(* IEC 61131-3 sources: daoli-st-library/DL_Device (part 39) *)

(* ---- FB_DL_HeatCoolZone.st ---- *)
(*==============================================================================
 * 组件名称 (Component)  : FB_DL_HeatCoolZone
 * 所属子库 (Sublibrary) : DL_Device
 * 当前版本 (Version)    : 1.0.0
 * 兼容性   (Platform)   : CODESYS 3.5 / TwinCAT 3 / 汇川 InoProShop / Machine Expert
 *                         仅依赖 Standard.library 语义与 DL_Algo 既有算法组件，
 *                         零厂商方言，零物理地址直写
 * 分类     (Category)   : 功能块（FUNCTION_BLOCK）· 加热/冷却温控区 · Level 1 DL_Device 开库件
 * 功能描述 (Function)   : 双通道（加热/冷却）温控区控制器，R4 算法族首个上层消费者。
 *                         控制链：FB_DL_PidController（含抗饱和，实例经引脚注入，
 *                         参数外置组态）→ 分程分配（Split-range，fSplitLow/High
 *                         可组态，非魔法数）→ FB_DL_PwmDutyController × 2（加热/
 *                         冷却 SSR 驱动）。断偶保护：传感器接口信号质量进入断线/
 *                         开路域时按 eBreakAction 切断对应通道并锁存 eSensorBreak
 *                         态（0003_0211），退出需 CmdReset 且质量恢复 eGood；
 *                         锁存期间双通道全断为最终安全态。设定值经 fTempMin/Max
 *                         钳位（信息级 0003_0101，不置故障）。本块零内嵌组态、
 *                         零魔法数，PID/PWM 全部实例经 IN_OUT 引脚注入。
 * 开源溯源 (Origin)     : 原创实现。分程控制与断偶安全方向为行业公知语义
 *                         （来源标签 lbp-device；断偶方向参考 NAMUR NE43 公开
 *                         标准），未复制任何厂商源码。PID/PWM 语义消费本库
 *                         DL_Algo 既有组件 FB_DL_PidController / FB_DL_PwmDutyController。
 * 本文件内含       : TYPE      E_DL_BreakAction（断偶动作方向枚举，归属 DL_Device）
 *                    FUNCTION_BLOCK FB_DL_HeatCoolZone IMPLEMENTS I_DL_TemperatureZone
 *                    （随附 METHOD ×3 与 PROPERTY GET ×5 实现体）
 * 依赖     (Depends)    : I_DL_TemperatureZone / E_DL_TempZoneState（同轮泳道交付
 *                          的 I_DL_TemperatureZone.st）；FB_DL_PidController、
 *                          FB_DL_PwmDutyController（DL_Algo v1.0.1+，实例注入）；
 *                          Standard.library：LIMIT / MIN / ABS。不引用库内任何
 *                          其他实现文件的具体逻辑。
 * 【规格偏离留档 / R11 Deviation register】
 *   D1 规格 §1.8 引脚表要求 fTempActual/fPowerOut/eState/bFault/uErrorId 五个
 *      「接口属性映射」成员同时作为 OUT 引脚暴露；IEC 61131-3 同一 POU 的变量
 *      与属性共享命名空间，同名变量与同名属性并存无法通过编译。按 R11 留档：
 *      该五成员以只读 PROPERTY 形式对外暴露（属性即输出引脚语义，接口成员逐一
 *      兑现），bHeaterOut/bCoolerOut 两个非接口成员保留 VAR_OUTPUT。
 *   D2（已闭环 / Closed）规格 §1.5 的 E_DL_SignalQuality / I_DL_AnalogSensor 为
 *      本块温度信号源契约。编码阶段宿主文件未入库，本文件曾就地声明副本；
 *      R5 注册收口阶段 I_DL_AnalogSensor.st（正式承载 E_DL_SignalQuality 枚举
 *      与 I_DL_AnalogSensor 接口）已随 DL_Device 开库交付，本文件重复副本已
 *      删除，改为引用该正式定义（IEC 同工程内 INTERFACE/ENUM 全局可见，与原
 *      D2 预设处置一致）。契约语义以 I_DL_AnalogSensor.st 为准（本块仅消费
 *      fValue 与 eQuality 两个成员）。
 *   D3 规格 §1.8「按 eBreakAction 切断对应通道并锁存」细化：eBreakAction 决定
 *      断偶瞬间立即切断的危险通道方向；锁存 eSensorBreak 期间双通道全断为最终
 *      安全态（锁存态不维持任何输出，安全侧选择）。
 *   D4 公约 0.6 示例码 16#0001_0001 属 DL_Base 段；按公约 0.7 段位分配（DL_Device
 *      族 16#0003_xxxx），本块参数钳位/对调修复统一置信息级 16#0003_0101。
 *   D5 新增故障/信息码顺延登记（无冲突）：16#0003_0212 非法状态兜底（故障级）、
 *      16#0003_0213 传感器接口引用未注入/无效（故障级）。
 * 故障码表（本块全部登记，0=无故障）：
 *   16#0003_0101【信息级】参数钳位/对调修复/设定值钳位提示，不置故障
 *   16#0003_0211【故障级】传感器断线/开路锁存，CmdReset + 质量恢复 eGood 方可清
 *   16#0003_0212【故障级】非法状态兜底（CASE ELSE 落点），CmdReset 可清
 *   16#0003_0213【故障级】温度传感器接口引用未注入/无效，CmdReset + 引脚有效方可清
 * 红线自检 (Redline)    : R1 ✓ 零全局变量表与外部变量引用 ｜ R2 ✓ 零物理 IO 地址直写
 *                         R3 ✓ 纯 IEC 61131-3 ｜ R4 ✓ 防除零+钳位+非有限值防御+浮点容差
 *                         R5 ✓ 全变量中英双语同行注释 ｜ R6 ✓ 六态 ENUM+CASE+ELSE 兜底
 *                         R7 ✓ 无直接定时器实例（PID/PWM 实例每拍无条件调用）
 * 修订历史 (Revision)   :
 *   2026-11-15  v1.0.0  首版入库 · Round 05 · 泳道 B · 契约出处 ROUND_PLAN_R5 §1.8
 *   2026-11-15  v1.0.0  R5 收口：删除就地重复的 E_DL_SignalQuality /
 *                       I_DL_AnalogSensor 声明，改引用 I_DL_AnalogSensor.st
 *                       正式定义（D2 闭环），功能与引脚零变更
 * 验收向量 (Acceptance) :
 *   V1 正常跃迁链：bEnable=TRUE → eHolding；fTempActual 低于设定 → eHeating；
 *      回到中性带 → eHolding；高于设定 → eCooling（fPowerOut 正负号随之翻转）
 *   V2 非法态兜底：强写内部状态为越界值 → CASE ELSE 落入 eFault（0003_0212）
 *   V3 中途跟踪脉冲（公约 0.1 必含）：闭环运行中 bTrack 单拍脉冲 + fTrackValue
 *      =30.0 → 本拍 PID 输出跟随 30.0，双通道占空比无扰重分配，无输出踢腿
 *   V4 断偶：eQuality=eWireBreakHigh → 按 eBreakAction 切断并锁存 eSensorBreak
 *      （0003_0211）；质量恢复 eGood + CmdReset → 回 eHolding（带无扰同步）
 *   V5 设定值钳位：fTempSetpoint=500 且 fTempMax=300 → 生效 300，0003_0101，
 *      故障位保持 FALSE（R21 信息级不置故障）
 *   V6 参数对调：fTempMin=300 > fTempMax=0 → 对调后继续计算，0003_0101
 *   V7 引脚无效：iTempSensor 未注入 → eFault（0003_0213），双通道切断
 *============================================================================*)

(*-----------------------------------------------------------------------------
 * 契约引用说明（R5 收口）: 本块温度信号源契约 E_DL_SignalQuality 与
 * I_DL_AnalogSensor 不在本文件就地声明，统一引用 DL_Device 正式定义文件
 * I_DL_AnalogSensor.st（枚举随宿主接口文件同文件发布，IEC 同工程内全局可见，
 * 留档见头注释 D2）。本块仅消费 fValue 与 eQuality 两个成员。
 *----------------------------------------------------------------------------*)

(*-----------------------------------------------------------------------------
 * 枚举: E_DL_BreakAction（归属 DL_Device，随 FB_DL_HeatCoolZone 同文件）
 * 含义: 断偶动作方向，按被控对象安全策略配置。
 *----------------------------------------------------------------------------*)
{attribute 'qualified_only'}
{attribute 'strict'}
TYPE E_DL_BreakAction :
(
    eHeatOff := 0,   // 断偶切断加热（Cut heating on break）：升温对象超温风险侧
    eCoolOff := 1    // 断偶切断冷却（Cut cooling on break）：骤冷风险对象（如防脆断工艺）侧
) UINT;
END_TYPE

(*==============================================================================
 * 功能块: FB_DL_HeatCoolZone IMPLEMENTS I_DL_TemperatureZone
 * 调用约定: 每个扫描周期无条件调用一次；PID/PWM 注入实例在本块主体每拍无条件
 *           调用（不在任何 IF/CASE 分支内部）；方法仅置请求标志，动作由主体执行。
 * 分程约定: PID 输出 [0..100 %]。输出低于 fSplitLow → 加热段（越低加热越强，
 *           配合 fKp 负值反作用）；高于 fSplitHigh → 冷却段（越高冷却越强）；
 *           两点之间为中性带（双通道全关，热平衡保持）。fSplitLow=0 时加热段
 *           跨度为零、加热通道自动禁用（防除零）；fSplitHigh=100 时同理禁用冷却。
 *============================================================================*)
FUNCTION_BLOCK FB_DL_HeatCoolZone IMPLEMENTS I_DL_TemperatureZone
VAR_INPUT
    fTempSetpoint   : REAL := 0.0;      // 目标温度（Setpoint）[°C]，经 fTempMin/Max 钳位后生效
    fTempMin        : REAL := 0.0;     // 设定值下边界（Setpoint lower bound）[°C]，默认 0.0
    fTempMax        : REAL := 300.0;   // 设定值上边界（Setpoint upper bound）[°C]，默认 300.0
    fSplitLow       : REAL := 50.0;    // 分程下切换点（Split-range low crossover）[%]，PID 输出低于此点进入加热段
    fSplitHigh      : REAL := 50.0;    // 分程上切换点（Split-range high crossover）[%]，PID 输出高于此点进入冷却段
    eBreakAction    : E_DL_BreakAction := E_DL_BreakAction.eHeatOff; // 断偶动作方向（Break action）：eHeatOff=切断加热 / eCoolOff=切断冷却
    bEnable         : BOOL := FALSE;   // 投运使能（Zone enable），与 CmdEnable 方法锁存值取与
    tSampleTime     : TIME := T#100MS; // 采样周期（Sample time），下传注入的 PID 与两路 PWM（公约 0.5）
    bTrack          : BOOL := FALSE;   // 跟踪使能（Track enable），TRUE 时本拍输出跟随 fTrackValue 无扰接管
    fTrackValue     : REAL := 0.0;     // 跟踪值（Track value）[-100..100 %]，与输出功率同量纲
END_VAR
VAR_IN_OUT
    iTempSensor     : I_DL_AnalogSensor;       // 温度信号源接口引用（Sensor interface reference），上层注入 FB_DL_AnalogTransmitter 实例
    fbPid           : FB_DL_PidController;     // 温度 PID 实例（Injected PID instance），增益/积分/限幅由调用方组态
    fbPwmHeat       : FB_DL_PwmDutyController; // 加热 SSR PWM 实例（Injected heat PWM），周期/最短脉冲由调用方组态
    fbPwmCool       : FB_DL_PwmDutyController; // 冷却 SSR PWM 实例（Injected cool PWM），周期/最短脉冲由调用方组态
END_VAR
VAR_OUTPUT
    bHeaterOut      : BOOL;            // 加热执行通道镜像（Heater channel mirror），等于加热 PWM 实例布尔输出
    bCoolerOut      : BOOL;            // 冷却执行通道镜像（Cooler channel mirror），等于冷却 PWM 实例布尔输出
END_VAR
VAR
    bInit           : BOOL := TRUE;    // 首扫标志（First-scan flag），首扫判据见段 1（公约 0.1 唯一合法范式）
    _eState         : E_DL_TempZoneState := E_DL_TempZoneState.eIdle; // 内部状态机步序（Internal zone state）
    _fTempActual    : REAL := 0.0;     // 实测温度快照（Actual temperature snapshot）[°C]，取自传感器接口
    _fPowerOut      : REAL := 0.0;     // 输出功率（Power output）[-100..100 %]，正=加热 / 负=冷却（R20 量纲与赋值式一致）
    _bFault         : BOOL := FALSE;   // 故障锁存标志（Fault latched），派生式：仅故障级状态置位，信息级不置位（R21）
    _uErrorId       : UDINT := 0;      // 故障/信息码（Error/info code），0=无；故障级进态写入、锁存保持
    _bCmdEnabled    : BOOL := TRUE;    // CmdEnable 方法锁存值（Method enable latch），默认投运（方法为可选入口）
    _fSetpointMethod: REAL := 0.0;     // SetSetpoint 方法锁存设定值（Method setpoint latch）[°C]，已按边界钳位
    _bUseMethodSp   : BOOL := FALSE;   // TRUE=方法设定值覆盖引脚设定值（Method setpoint override）
    _bSyncReq       : BOOL := FALSE;   // 跃迁无扰同步请求（Bumpless sync request），置位后下一拍 PID 跟踪当前功率
    _bTrackActive   : BOOL := FALSE;   // 本拍处于外部跟踪（External track active this scan），由段 1 判据得出
    _fPowerOutLast  : REAL := 0.0;     // 上一拍输出功率（Last power output）[-100..100 %]，跃迁同步的跟踪源
    _fTempMinEff    : REAL := 0.0;     // 修复后设定值下边界（Repaired lower bound）[°C]
    _fTempMaxEff    : REAL := 300.0;   // 修复后设定值上边界（Repaired upper bound）[°C]
    _fSplitLowEff   : REAL := 50.0;    // 修复后分程下切换点（Repaired low crossover）[%]
    _fSplitHighEff  : REAL := 50.0;    // 修复后分程上切换点（Repaired high crossover）[%]
    _fSpEff         : REAL := 0.0;     // 有效设定值（Effective setpoint）[°C]，来源仲裁 + 钳位后
    _fTrackSrc      : REAL := 0.0;     // 本拍跟踪源（Track source this scan）[-100..100 %]
    _fPidOut        : REAL := 0.0;     // PID 输出快照（PID output snapshot）[0..100 %]
    _fHeatDuty      : REAL := 0.0;     // 加热通道占空比（Heater duty）[0..100 %]
    _fCoolDuty      : REAL := 0.0;     // 冷却通道占空比（Cooler duty）[0..100 %]
    _fSpTmp         : REAL := 0.0;     // 参数对调临时变量（Swap temporary）[°C 或 %]
    _bRefOk         : BOOL := FALSE;   // 传感器接口引用有效标志（Sensor reference valid）
    _bSensorBad     : BOOL := FALSE;   // 传感器断线/开路标志（Sensor break flag），含非有限值防御归入
    _bInfoClamp     : BOOL := FALSE;   // 本拍发生钳位/对调修复（Info-level clamp occurred）
    _bRunPre        : BOOL := FALSE;   // CASE 前运行态判定（Pre-CASE running flag），PID 使能源
    _bZoneRun       : BOOL := FALSE;   // CASE 后运行态判定（Post-CASE running flag），PWM 使能源
    _bReqEnable     : BOOL := FALSE;   // CmdEnable 请求挂起（Enable request pending）
    _bValEnable     : BOOL := FALSE;   // CmdEnable 请求值（Enable request value）
    _bReqReset      : BOOL := FALSE;   // CmdReset 请求挂起（Reset request pending）
    _bReqSetSp      : BOOL := FALSE;   // SetSetpoint 请求挂起（Setpoint request pending）
    _fReqSetSp      : REAL := 0.0;     // SetSetpoint 请求原始值（Raw setpoint request）[°C]
    _eQuality       : E_DL_SignalQuality := E_DL_SignalQuality.eGood; // 传感器信号质量快照（Quality snapshot）
END_VAR
VAR CONSTANT
    DL_ZONE_POWER_TOL : REAL := 0.01;   // 热平衡零功率判定容差（Power tolerance）[%]，浮点容差红线，状态判稳阈值
    DL_ZONE_SPAN_EPS  : REAL := 1.0E-6; // 分程跨度防除零判据（Span epsilon）[%]，低于此值通道禁用
END_VAR

METHOD SetSetpoint : BOOL
VAR_INPUT
    fTemp : REAL;                        // 目标温度（Target temperature）[°C]，非有限值拒绝
END_VAR
// 返回合法性：非有限值一律拒绝（公约 0.8 判式），合法值锁存待主体钳位生效
IF fTemp <> fTemp THEN
    SetSetpoint := FALSE;                // 非有限值拒绝
ELSE
    _fReqSetSp := fTemp;                 // 请求原始值 [°C]
    _bReqSetSp := TRUE;                  // 置单发标志，主体段 2/段 3 落实
    SetSetpoint := TRUE;                 // 受理成功
END_IF

    END_METHOD

METHOD CmdEnable
VAR_INPUT
    bOn : BOOL;                          // TRUE=投运（Commission on），FALSE=退出并切断双通道
END_VAR
_bReqEnable := TRUE;                     // 置请求标志
_bValEnable := bOn;                      // 请求值随行

    END_METHOD

METHOD CmdReset : BOOL
// 返回当前是否可复位：断偶锁存态要求信号质量快照已恢复 eGood（规格 §1.8 退出条件）
_bReqReset := TRUE;                      // 置请求标志，主体段 7 各态消费
IF _eState = E_DL_TempZoneState.eSensorBreak THEN
    IF _bRefOk AND (_eQuality = E_DL_SignalQuality.eGood) AND (NOT _bSensorBad) THEN
        CmdReset := TRUE;                // 质量已恢复，可复位
    ELSE
        CmdReset := FALSE;               // 仍在断线域，拒绝复位
    END_IF
ELSE
    CmdReset := TRUE;                    // 非断偶态一律受理
END_IF

// =============================================================================
// 属性实现区（PROPERTY GET ×5，接口契约逐字兑现；偏离 D1：属性即输出引脚语义）
// =============================================================================

    END_METHOD

// -----------------------------------------------------------------------------
// 段 1｜首扫与跟踪同步（公约 0.1 / R19 唯一合法范式：跟踪项在前、首扫项取反在后，
//       禁止两项顺序颠倒的反式写法；验收向量 V3 覆盖运行中途跟踪脉冲）
// -----------------------------------------------------------------------------
IF bTrack OR (NOT bInit) THEN
    _fPowerOutLast := 0.0;               // 首扫/外部跟踪：历史功率清零，杜绝接管瞬间踢腿 [±100 %]
    _bTrackActive  := TRUE;              // 本拍输出跟随外部跟踪值 fTrackValue
    bInit          := TRUE;              // 首扫完成置位
ELSE
    _bTrackActive  := FALSE;             // 正常闭环拍，跟踪源取内部历史功率
END_IF

// -----------------------------------------------------------------------------
// 段 2｜方法请求消费（方法内只置标志，动作在本周期落实——跨周期动作不驻留方法）
// -----------------------------------------------------------------------------
IF _bReqEnable THEN
    _bCmdEnabled := _bValEnable;         // 投/退锁存值更新
    _bReqEnable  := FALSE;               // 单发消费
END_IF
IF _bReqSetSp THEN
    _fSetpointMethod := _fReqSetSp;      // 方法设定值锁存 [°C]，边界钳位在段 3 统一进行
    _bUseMethodSp    := TRUE;            // 方法设定值覆盖引脚设定值
    _bReqSetSp       := FALSE;           // 单发消费
END_IF
IF NOT ( (_eState = E_DL_TempZoneState.eSensorBreak) OR (_eState = E_DL_TempZoneState.eFault) ) THEN
    _bReqReset := FALSE;                 // 非锁存态下的复位请求立即作废，防陈旧请求迟到生效
END_IF

// -----------------------------------------------------------------------------
// 段 3｜参数修复（公约 0.6 对调自修复 + 公约 0.8 非有限值防御；信息级 0003_0101
//       只进 uErrorId 不置故障，R21；偏离 D4：段位按公约 0.7 归 DL_Device 族）
// -----------------------------------------------------------------------------
_bInfoClamp := FALSE;
IF fTempMin <> fTempMin THEN             // NaN 恒不等于自身（公约 0.8 指定判式）
    _fTempMinEff := 0.0;                 // 非有限值回退默认下边界 [°C]
    _bInfoClamp  := TRUE;
ELSE
    _fTempMinEff := fTempMin;            // 直接采纳 [°C]
END_IF
IF fTempMax <> fTempMax THEN
    _fTempMaxEff := 300.0;               // 非有限值回退默认上边界 [°C]
    _bInfoClamp  := TRUE;
ELSE
    _fTempMaxEff := fTempMax;            // 直接采纳 [°C]
END_IF
IF _fTempMinEff > _fTempMaxEff THEN      // 边界对调自修复（公约 0.6）：修复后继续计算，不中断
    _fSpTmp       := _fTempMinEff;
    _fTempMinEff  := _fTempMaxEff;
    _fTempMaxEff  := _fSpTmp;
    _bInfoClamp   := TRUE;
END_IF

IF fSplitLow <> fSplitLow THEN
    _fSplitLowEff := 50.0;               // 非有限值回退对称默认 [%]
    _bInfoClamp   := TRUE;
ELSE
    _fSplitLowEff := fSplitLow;          // 直接采纳 [%]
END_IF
IF fSplitHigh <> fSplitHigh THEN
    _fSplitHighEff := 50.0;              // 非有限值回退对称默认 [%]
    _bInfoClamp    := TRUE;
ELSE
    _fSplitHighEff := fSplitHigh;        // 直接采纳 [%]
END_IF
IF _fSplitLowEff < 0.0 THEN
    _fSplitLowEff := 0.0;                // 钳到分程域下限 [%]（此时加热段跨度为零，加热禁用）
    _bInfoClamp   := TRUE;
END_IF
IF _fSplitLowEff > 100.0 THEN
    _fSplitLowEff := 100.0;              // 钳到分程域上限 [%]
    _bInfoClamp   := TRUE;
END_IF
IF _fSplitHighEff < 0.0 THEN
    _fSplitHighEff := 0.0;               // 钳到分程域下限 [%]
    _bInfoClamp    := TRUE;
END_IF
IF _fSplitHighEff > 100.0 THEN
    _fSplitHighEff := 100.0;             // 钳到分程域上限 [%]（此时冷却段跨度为零，冷却禁用）
    _bInfoClamp    := TRUE;
END_IF
IF _fSplitLowEff > _fSplitHighEff THEN   // 分程点对调自修复（公约 0.6）
    _fSpTmp        := _fSplitLowEff;
    _fSplitLowEff  := _fSplitHighEff;
    _fSplitHighEff := _fSpTmp;
    _bInfoClamp    := TRUE;
END_IF

// 设定值来源仲裁：方法锁存值优先，否则取引脚连续值
IF _bUseMethodSp THEN
    _fSpEff := _fSetpointMethod;         // 方法通道 [°C]
ELSE
    _fSpEff := fTempSetpoint;            // 引脚通道 [°C]
END_IF
IF _fSpEff <> _fSpEff THEN
    _fSpEff     := _fTempMinEff;         // 非有限设定值回退下边界（安全侧低温待机）[°C]
    _bInfoClamp := TRUE;
END_IF
IF (_fSpEff < _fTempMinEff) OR (_fSpEff > _fTempMaxEff) THEN
    _fSpEff     := LIMIT(_fTempMinEff, _fSpEff, _fTempMaxEff);  // 设定值钳位（规格 §1.8 设计点，信息级 0003_0101）
    _bInfoClamp := TRUE;
END_IF

// -----------------------------------------------------------------------------
// 段 4｜传感器采集与有效性判定（接口引用检查 + 质量域 + 非有限值防御）
// -----------------------------------------------------------------------------
_bRefOk     := FALSE;
_bSensorBad := FALSE;
_eQuality   := E_DL_SignalQuality.eGood;
IF iTempSensor <> 0 THEN                 // 接口引用有效性检查（未注入防御）
    _bRefOk     := TRUE;
    _fTempActual := iTempSensor.fValue;  // 工程量实测值 [°C]，契约保证 NaN 防御后输出
    _eQuality    := iTempSensor.eQuality;
    IF _fTempActual <> _fTempActual THEN
        _bSensorBad := TRUE;             // 非有限值防御：NaN 按断线域处理（公约 0.8 判式）
    ELSIF (_eQuality = E_DL_SignalQuality.eWireBreakLow)
       OR (_eQuality = E_DL_SignalQuality.eWireBreakHigh)
       OR (_eQuality = E_DL_SignalQuality.eOpenLoop) THEN
        _bSensorBad := TRUE;             // NE43 断线/开路域（规格 §1.8 断偶保护集合）
    END_IF
END_IF

// -----------------------------------------------------------------------------
// 段 5｜运行态预判定与注入 PID 无条件调用（R7 精神：实例调用不在 IF/CASE 分支内）
// -----------------------------------------------------------------------------
_bRunPre := (_eState = E_DL_TempZoneState.eHolding)
         OR (_eState = E_DL_TempZoneState.eHeating)
         OR (_eState = E_DL_TempZoneState.eCooling);
IF _bTrackActive THEN
    _fTrackSrc := fTrackValue;           // 外部跟踪源 [-100..100 %]
ELSE
    _fTrackSrc := _fPowerOutLast;        // 跃迁同步源 = 上一拍实际输出功率 [-100..100 %]
END_IF
fbPid(
    bEnable     := _bRunPre AND _bRefOk AND (NOT _bSensorBad),  // 断偶/无引用时冻结 PID（输出回下限）
    bManual     := FALSE,                // 温控区纯自动模式，手动路径不由本块开放
    fSetpoint   := _fSpEff,              // 有效设定值 [°C]
    fActual     := _fTempActual,         // 实测温度 [°C]
    tSampleTime := tSampleTime,          // 采样周期下传（公约 0.5）
    bTrack      := _bTrackActive OR _bSyncReq,  // 外部跟踪或跃迁无扰同步（电平，一拍）
    fTrackValue := _fTrackSrc            // 跟踪值 [-100..100 %]
);
_bSyncReq := FALSE;                      // 同步请求单发消费（段 7 跃迁时重新置位）

// -----------------------------------------------------------------------------
// 段 6｜分程分配（热平衡计算，防除零：跨度不足的通道自动禁用，R4 红线）
// -----------------------------------------------------------------------------
IF _bRunPre AND _bRefOk AND (NOT _bSensorBad) THEN
    _fPidOut := fbPid.fOut;              // PID 输出 [0..100 %]，量程由调用方组态
    IF _fPidOut < _fSplitLowEff THEN
        // 加热段：输出越低于下切换点，加热越强（配合 fKp 负值反作用惯例）
        IF _fSplitLowEff > DL_ZONE_SPAN_EPS THEN
            _fHeatDuty := LIMIT(0.0, (_fSplitLowEff - _fPidOut) / _fSplitLowEff * 100.0, 100.0); // 加热占空比 [0..100 %]
        ELSE
            _fHeatDuty := 0.0;           // 加热段跨度为零，通道禁用（防除零）
        END_IF
        _fCoolDuty := 0.0;               // 加热段冷却通道必关 [0..100 %]
    ELSIF _fPidOut > _fSplitHighEff THEN
        // 冷却段：输出越高于上切换点，冷却越强
        IF (100.0 - _fSplitHighEff) > DL_ZONE_SPAN_EPS THEN
            _fCoolDuty := LIMIT(0.0, (_fPidOut - _fSplitHighEff) / (100.0 - _fSplitHighEff) * 100.0, 100.0); // 冷却占空比 [0..100 %]
        ELSE
            _fCoolDuty := 0.0;           // 冷却段跨度为零，通道禁用（防除零）
        END_IF
        _fHeatDuty := 0.0;               // 冷却段加热通道必关 [0..100 %]
    ELSE
        _fHeatDuty := 0.0;               // 中性带：双通道全关，热平衡保持 [0..100 %]
        _fCoolDuty := 0.0;               // 中性带 [0..100 %]
    END_IF
ELSE
    _fPidOut   := 0.0;                   // 非运行拍 PID 输出按 0 [%] 处理
    _fHeatDuty := 0.0;                   // 非运行拍加热占空比清零 [0..100 %]
    _fCoolDuty := 0.0;                   // 非运行拍冷却占空比清零 [0..100 %]
END_IF
_fPowerOut := _fHeatDuty - _fCoolDuty;   // 输出功率 [-100..100 %]，正=加热/负=冷却（R20 量纲与赋值式一致）

// -----------------------------------------------------------------------------
// 段 7｜状态机（ENUM + CASE + ELSE 兜底；断偶/非法态/无引用均为锁存，R15 仅复位可清）
// -----------------------------------------------------------------------------
CASE _eState OF

    E_DL_TempZoneState.eIdle:            // 空闲：双通道切断（PWM 使能在段 8 落实）
        IF _bRefOk AND (NOT _bSensorBad) AND bEnable AND _bCmdEnabled THEN
            _bSyncReq := TRUE;           // 投运首拍无扰同步，PID 跟踪当前功率 0 [%]
            _eState   := E_DL_TempZoneState.eHolding;
        END_IF

    E_DL_TempZoneState.eHolding:         // 保温：双通道处于热平衡容差带
        IF NOT (bEnable AND _bCmdEnabled) THEN
            _eState := E_DL_TempZoneState.eIdle;
        ELSIF NOT _bRefOk THEN
            _uErrorId := 16#0003_0213;   // 接口引用未注入/无效（故障级锁存）
            _eState   := E_DL_TempZoneState.eFault;
        ELSIF _bSensorBad THEN
            _uErrorId := 16#0003_0211;   // 断偶锁存（故障级；eBreakAction 切断方向语义见偏离 D3）
            _eState   := E_DL_TempZoneState.eSensorBreak;
        ELSIF _fPowerOut > DL_ZONE_POWER_TOL THEN
            _eState := E_DL_TempZoneState.eHeating;
        ELSIF _fPowerOut < -DL_ZONE_POWER_TOL THEN
            _eState := E_DL_TempZoneState.eCooling;
        END_IF

    E_DL_TempZoneState.eHeating:         // 加热中
        IF NOT (bEnable AND _bCmdEnabled) THEN
            _eState := E_DL_TempZoneState.eIdle;
        ELSIF NOT _bRefOk THEN
            _uErrorId := 16#0003_0213;   // 接口引用未注入/无效
            _eState   := E_DL_TempZoneState.eFault;
        ELSIF _bSensorBad THEN
            _uErrorId := 16#0003_0211;   // 断偶锁存
            _eState   := E_DL_TempZoneState.eSensorBreak;
        ELSIF _fPowerOut < -DL_ZONE_POWER_TOL THEN
            _eState := E_DL_TempZoneState.eCooling;
        ELSIF ABS(_fPowerOut) <= DL_ZONE_POWER_TOL THEN
            _eState := E_DL_TempZoneState.eHolding;   // 回到热平衡带（浮点容差红线）
        END_IF

    E_DL_TempZoneState.eCooling:         // 冷却中
        IF NOT (bEnable AND _bCmdEnabled) THEN
            _eState := E_DL_TempZoneState.eIdle;
        ELSIF NOT _bRefOk THEN
            _uErrorId := 16#0003_0213;   // 接口引用未注入/无效
            _eState   := E_DL_TempZoneState.eFault;
        ELSIF _bSensorBad THEN
            _uErrorId := 16#0003_0211;   // 断偶锁存
            _eState   := E_DL_TempZoneState.eSensorBreak;
        ELSIF _fPowerOut > DL_ZONE_POWER_TOL THEN
            _eState := E_DL_TempZoneState.eHeating;
        ELSIF ABS(_fPowerOut) <= DL_ZONE_POWER_TOL THEN
            _eState := E_DL_TempZoneState.eHolding;   // 回到热平衡带
        END_IF

    E_DL_TempZoneState.eSensorBreak:     // 断偶锁存：双通道全断（安全终态，偏离 D3）
        IF _bReqReset AND _bRefOk AND (_eQuality = E_DL_SignalQuality.eGood)
           AND (NOT _bSensorBad) AND bEnable AND _bCmdEnabled THEN
            _bReqReset := FALSE;         // 复位请求消费
            _bSyncReq  := TRUE;          // 复位回投无扰同步
            _eState    := E_DL_TempZoneState.eHolding;
        END_IF

    E_DL_TempZoneState.eFault:           // 故障兜底：双通道全断
        IF _bReqReset AND _bRefOk THEN
            _bReqReset := FALSE;         // 复位请求消费（引用已恢复有效）
            _bSyncReq  := TRUE;          // 复位回投无扰同步
            _eState    := E_DL_TempZoneState.eHolding;
        END_IF

    ELSE                                 // 非法状态兜底拦截（R6 红线）
        _uErrorId := 16#0003_0212;       // 非法状态（故障级锁存）
        _eState   := E_DL_TempZoneState.eFault;
END_CASE

// -----------------------------------------------------------------------------
// 段 8｜注入 PWM 无条件调用与输出镜像（R7 精神：实例调用不在 IF/CASE 分支内）
// -----------------------------------------------------------------------------
_bZoneRun := (_eState = E_DL_TempZoneState.eHolding)
          OR (_eState = E_DL_TempZoneState.eHeating)
          OR (_eState = E_DL_TempZoneState.eCooling);
fbPwmHeat(
    bEnable     := _bZoneRun,            // 锁存态/空闲态强制关断
    fDuty       := _fHeatDuty,           // 加热占空比 [0..100 %]
    tSampleTime := tSampleTime,          // 采样周期下传（公约 0.5）
    bInvert     := FALSE                 // 正相输出
);
fbPwmCool(
    bEnable     := _bZoneRun,            // 锁存态/空闲态强制关断
    fDuty       := _fCoolDuty,           // 冷却占空比 [0..100 %]
    tSampleTime := tSampleTime,          // 采样周期下传（公约 0.5）
    bInvert     := FALSE                 // 正相输出
);
bHeaterOut := fbPwmHeat.bPwmOut;         // 加热通道镜像 = 注入 PWM 布尔输出
bCoolerOut := fbPwmCool.bPwmOut;         // 冷却通道镜像 = 注入 PWM 布尔输出

// -----------------------------------------------------------------------------
// 段 9｜故障派生（R21：bFault 为显式排除信息级码的派生式）与历史存档
// -----------------------------------------------------------------------------
_bFault := (_eState = E_DL_TempZoneState.eSensorBreak)
        OR (_eState = E_DL_TempZoneState.eFault);       // 仅故障级状态置位，0003_0101 不置位
IF _eState = E_DL_TempZoneState.eSensorBreak THEN
    _uErrorId := 16#0003_0211;           // 断偶锁存码逐拍保持，直至复位
ELSIF _eState <> E_DL_TempZoneState.eFault THEN
    IF _bInfoClamp THEN
        _uErrorId := 16#0003_0101;       // 信息级：钳位/对调修复提示，不置故障（R19）
    ELSE
        _uErrorId := 16#0000_0000;       // 无故障无提示
    END_IF
END_IF
// eFault 态不重写 _uErrorId：保持进态时写入的 0212/0213，锁存至复位（R15）
_fPowerOutLast := _fPowerOut;            // 存档本拍功率，供下一拍跃迁同步跟踪 [-100..100 %]

// =============================================================================
// 方法实现区（METHOD，共 3 个，接口契约逐字兑现；非阻塞单发语义）
// =============================================================================

PROPERTY fTempActual : REAL
fTempActual := _fTempActual;             // 实测温度 [°C]

PROPERTY fPowerOut : REAL
fPowerOut := _fPowerOut;                 // 输出功率 [-100..100 %]，正=加热/负=冷却

PROPERTY eState : E_DL_TempZoneState
eState := _eState;                       // 当前温控区状态

PROPERTY bFault : BOOL
bFault := _bFault;                       // 故障锁存标志（派生式，信息级不置位）

PROPERTY uErrorId : UDINT
uErrorId := _uErrorId;                   // 末次故障/信息码

END_FUNCTION_BLOCK

(* ---- FB_DL_IonFanInterlock.st ---- *)
(*
  ==================================================================
  组件名 Component  : FB_DL_IonFanInterlock
  分类   Category   : DL_Device
  前缀   Naming     : FB_DL_ ｜ b/n/u/f/t/e/st 类型前缀制（R265）
  码位   Code ID    : 16#0003_0717 / 0718 / 0719 / 071A（故障级）｜ 16#0003_071B / 071C（信息级）
  版本   Version    : 1.0.1
  复杂度 Complexity  : 中
  功能   Purpose    : 离子风机「运行反馈 + 风速下限 + 平衡电压」三判据合取，输出下游设备的
                      许可位（半导体 / 锂电装配段 ESD 防护联锁）。
  开源溯源 Origin    : IEC 61131-3 标准语义的道莅防御性实现（clean-room，无第三方代码行）；
                      NE107 诊断分级口径（Failure / OutOfSpec）为公开标准的分类借鉴，
                      零代码复制；闸门、迟滞、非对称许可与码位 100% 自有。
  许可证 License    : MIT
  参考   Reference  : IEC 61131-3:2013 §6.6 算术运算符；ISA-107 / NE107 诊断分级语义
                      （分类借鉴）；离子风机效能判据的公开 ESD 工程口径
  平台   Platform   : 纯 IEC 61131-3（TON / CASE / 四则 / 比较），三平台通用
  依赖   Depends    : 仅 Standard.library（TON 属标准定时器）
  分工声明 Split     : FB_DL_VacIonizerBalance 为平衡电压测量 / 标定属主（本件只消费其
                      结果或现场模拟量，绝不重算平衡）；FB_DL_AirShowerInterlockSeq 为
                      风淋门物流联锁；FB_DL_EsdGroundMonitor 为接地连续性；本件为离子风机
                      效能联锁，四件边界写死（R216 双向互引，选型见 MANUAL_DL_Device）。
  归属 Ownership     : E_DL_IonFanPhase 属主为本文件（全库唯一定义，R264）；引用件只引用
                      不重声明。
  ------------------------------------------------------------------
  边界 Boundary     :
                      一 许可发放非对称（本件核心安全口径，写死）：许可发放可延迟（须三判据
                         同时满足并持续 tConfirm），许可撤除零延时（任一判据失效当拍即
                         bPermit = FALSE）——TON 只作用于「发放」，撤除不经过任何定时器；
                      二 首拍 _bInit → bPermit := FALSE（出厂默认 F，禁首拍误许可）；bEnable
                         由 F 转 T 且判据已满足时仍须完整走完 tConfirm（禁跳过确认窗）；
                      三 判据迟滞（fHystPct）两方向分别定义，禁合成单一阈值：
                         风速下限：低于 fSpeedMin × (1 − h%) 置警、高于 fSpeedMin × (1 + h%) 复原；
                         平衡上限：高于 fBalanceLimV 置警、低于 fBalanceLimV × (1 − h%) 复原
                         （方向性证明：限 5 V 时 6 V 置警、回落 4.9 V 仍报警，因 4.9 > 4.75）；
                      四 非有限输入（fAirSpeed / fBalanceV 为 NaN 或 ±Inf）一律保守判不满足并
                         置对应故障码，区分「测点坏」与「真超标」（前者 bValid = FALSE +
                         独立码，后者为信息级 OutOfSpec）；
                      五 组态域闸：fSpeedMin ≤ 0、fBalanceLimV ≤ 0、tConfirm ≤ T#0S、fHystPct < 0
                         或任一限值非有限 → 组态故障码 + bPermit := FALSE；
                      六 状态机 ENUM + CASE 必带 ELSE；ELSE 落 eAlarm 并清许可（禁静默）；
                         TON 段 0 无条件刷新（禁入分支，R7）；TON IN 串组态闸与使能；
                      七 故障码逐拍重算不锁存（本件无 bReset 引脚，R152 解除路径自证：
                         解除路径 = 修正组态 / 恢复测点，两条恒可达）；首因保序由判据顺序保证；
                      八 bEnable = FALSE（v1.0.1 返修 R63 · 修 R62-D3：按 R300 取「实现串
                         bEnable」口径）：bPermit := FALSE、三报警位（bAlarmSpeed /
                         bAlarmBalance / bAlarmFan）全部串 bEnable 归零、bError 串
                         bEnable 归零、eErr 归零不发码——失能相不再外显 Failure 级
                         假故障（R191 名实双出口：信号出口与状态出口同源）；
                      九 段序（v1.0.1 顺带消除 R62-D6 轻项）：组态域闸先行（段 0），
                         段 1 判据与 tonConfirm 使用本拍组态位，不再引用上一拍值。
  错误码 Codes      :
    16#0003_0717【故障级】组态非法（fSpeedMin ≤ 0 / fBalanceLimV ≤ 0 / tConfirm ≤ 0 / fHystPct < 0 / 限值非有限）
    16#0003_0718【故障级】风机运行反馈丧失（Failure 级，零延时撤销许可）
    16#0003_0719【故障级】风速测点非有限（NaN 或 ±Inf，测点坏而非真超标）
    16#0003_071A【故障级】平衡电压测点非有限（NaN 或 ±Inf，测点坏而非真超标）
    16#0003_071B【信息级】风速低于下限（OutOfSpec，bAlarmSpeed = TRUE）
    16#0003_071C【信息级】平衡电压超限（OutOfSpec，bAlarmBalance = TRUE）
  码位反证 Note     :
    0719 / 071A 与 071B / 071C 必须分开：测点坏的处置人是仪表工（换探头 / 查接线），
    真超标的处置人是工艺工程师（调风机 / 查高压发生器），而两者的 bPermit 与报警位组合
    完全相同（bPermit = FALSE、报警位 TRUE），仅靠输出无法区分，故各自独立码（R90）。
  验收 Acceptance   :
    算法已证（脚本）：未跑 ｜ 编译器已证（三平台）：未跑
    V1 三判据全满足并持续 tConfirm → bPermit = TRUE、eState = ePermit
    V2 tConfirm 未到即撤除 → 全程 bPermit = FALSE
    V3 许可态下 bFanRun 掉电 → 同拍 bPermit = FALSE + bAlarmFan（零延时撤除向量）
    V4 fAirSpeed = NaN → bPermit = FALSE + 码 0719 + bValid = FALSE
    V5 fSpeedMin = 0 → 码 0717 + bPermit = FALSE
    V6 风速在 fSpeedMin 上下抖动 3%（小于迟滞 5%）→ 判据不反复跳
    V7 平衡电压 +6 V（限 5 V）→ bAlarmBalance = TRUE、bPermit = FALSE；回落 4.9 V 仍报警
    V8 首拍 → bPermit = FALSE
    V9 bEnable 由 F 转 T 且判据已满足 → 仍需完整 tConfirm
  修订记录 Revision  :
    2026-11-21  v1.0.0  R62 首版（批 4 · 序号 11；承接 ROADMAP R56-1086 半勾项）
    2026-11-21  v1.0.1  R63 返修 R3（R62-D3 中）：出口三报警位与 bError 全部串 bEnable，
                        失能相不再外显 Failure 级假故障；eErr 回放失能相归零；
                        顺带消除 R62-D6（轻）：组态闸提为段 0 先行，tonConfirm 改用本拍组态位
  ==================================================================
*)
TYPE E_DL_IonFanPhase :
(
    eIdle   := 0,  // 空闲：未使能或已失能 / idle, disabled
    eWarmup := 10, // 确认中：三判据满足并正在计时 tConfirm / confirming, the three criteria hold while the timer runs
    ePermit := 20, // 已许可：下游允许运行 / permitted, the downstream may run
    eAlarm  := 30  // 判据失效报警：许可已撤除 / an alarm, the permit has been withdrawn
);
END_TYPE

FUNCTION_BLOCK FB_DL_IonFanInterlock
VAR_INPUT
    bEnable       : BOOL := TRUE;        // 使能，FALSE 时清许可并回空闲（边界八）/ the enable, false clears the permit and returns to idle
    bFanRun       : BOOL := FALSE;       // 风机运行反馈 [-] / the fan running feedback
    fAirSpeed     : LREAL := 0.0;        // 出风速度 [米每秒]，必须有限 / the air speed, must be finite
    fSpeedMin     : LREAL := 0.5;        // 风速下限 [米每秒]，须 > 0 / the air speed floor, must be positive
    fBalanceV     : LREAL := 0.0;        // 离子平衡电压实测 [伏]，必须有限 / the measured balance voltage, must be finite
    fBalanceLimV  : LREAL := 5.0;        // 平衡电压绝对上限 [伏]，须 > 0 / the balance voltage absolute limit, must be positive
    tConfirm      : TIME := T#3S;        // 判据持续确认窗 [毫秒]，须 > 0 / the confirmation window, must be positive
    fHystPct      : LREAL := 5.0;        // 判据迟滞 [%]，须 ≥ 0 / the criterion hysteresis in percent, non negative
END_VAR
VAR_OUTPUT
    bPermit       : BOOL := FALSE;            // 下游允许运行（安全侧默认 FALSE，边界一）/ the downstream permit, safe side default false
    bAlarmSpeed   : BOOL := FALSE;            // 风速判据报警（OutOfSpec 级）[-] / the air speed alarm
    bAlarmBalance : BOOL := FALSE;            // 平衡电压判据报警（OutOfSpec 级）[-] / the balance voltage alarm
    bAlarmFan     : BOOL := FALSE;            // 风机运行反馈丧失报警（Failure 级）[-] / the fan feedback loss alarm
    eState        : E_DL_IonFanPhase;         // 状态机出口 [状态] / the state machine outlet
    bValid        : BOOL := FALSE;            // 测量可用（无测点故障与组态故障）[-] / the measurement is usable
    eErr          : UDINT := 16#0000_0000;    // 错误码，0 = 正常 / the error code, zero is ok
    bError        : BOOL := FALSE;            // 故障标志（故障级码同拍置位，R45 配对）/ the fault flag raised with a fault level code
END_VAR
VAR
    _bInit      : BOOL := FALSE;                        // 首拍初始化标志（R310）/ the first scan flag
    _eState     : E_DL_IonFanPhase := E_DL_IonFanPhase.eIdle; // 内部状态寄存器 / the internal state register
    _bFanOk     : BOOL := FALSE;                        // 风机运行判据（逐拍重算）/ the fan criterion
    _bSpeedOk   : BOOL := FALSE;                        // 风速判据（带迟滞，逐拍重算）/ the air speed criterion with hysteresis
    _bBalOk     : BOOL := FALSE;                        // 平衡电压判据（带迟滞，逐拍重算）/ the balance criterion with hysteresis
    _bAllOk     : BOOL := FALSE;                        // 三判据合取（逐拍重算）/ the conjunction of the three criteria
    _bAlmSpd    : BOOL := FALSE;                        // 风速报警迟滞状态（跨拍保持）/ the air speed alarm hysteresis state
    _bAlmBal    : BOOL := FALSE;                        // 平衡电压报警迟滞状态（跨拍保持）/ the balance alarm hysteresis state
    _bFinSpd    : BOOL := FALSE;                        // 风速测点有限标记（逐拍重算）/ the air speed finiteness flag
    _bFinBal    : BOOL := FALSE;                        // 平衡测点有限标记（逐拍重算）/ the balance finiteness flag
    _bCfgBad    : BOOL := FALSE;                        // 组态非法标记（逐拍重算）/ the configuration fault flag
    _fSpdTrip   : LREAL := 0.0;                         // 风速置警阈值 [米每秒] / the air speed trip threshold
    _fSpdRele   : LREAL := 0.0;                         // 风速复原阈值 [米每秒] / the air speed release threshold
    _fBalTrip   : LREAL := 0.0;                         // 平衡置警阈值（绝对值）[伏] / the balance trip threshold
    _fBalRele   : LREAL := 0.0;                         // 平衡复原阈值（绝对值）[伏] / the balance release threshold
    _fBalAbs    : LREAL := 0.0;                         // 平衡电压绝对值 [伏] / the absolute balance voltage
    _fPctScale  : LREAL := 0.0;                         // 迟滞百分比换算中间量 [−] / the hysteresis percentage intermediate
    tonConfirm  : TON;                                  // 判据持续确认定时器，段 0 无条件刷新 / the confirmation timer refreshed unconditionally
END_VAR  // R64 结构补齐：VAR 段缺失的 END_VAR（门禁机械修复）
VAR CONSTANT
    DL_IFI_ZERO  : LREAL := 0.0;   // 实数零常量 [工程单位] / the real zero constant
    DL_IFI_HUND  : LREAL := 100.0; // 百分比换算系数 [%] / the percentage scaling factor
    DL_IFI_TIME0 : TIME := T#0S;   // 时间零常量 [毫秒] / the time zero constant
END_VAR

// 段 0｜组态域闸先行（v1.0.1 修 R62-D6：tonConfirm 与判据段改用本拍组态位，禁用上一拍值，R272 全量点名）/ segment 0, the configuration gate runs first
_bCfgBad := (fSpeedMin <> fSpeedMin) OR ((fSpeedMin - fSpeedMin) <> (fSpeedMin - fSpeedMin)) OR (fSpeedMin <= DL_IFI_ZERO)
         OR (fBalanceLimV <> fBalanceLimV) OR ((fBalanceLimV - fBalanceLimV) <> (fBalanceLimV - fBalanceLimV)) OR (fBalanceLimV <= DL_IFI_ZERO)
         OR (fHystPct <> fHystPct) OR ((fHystPct - fHystPct) <> (fHystPct - fHystPct)) OR (fHystPct < DL_IFI_ZERO)
         OR (tConfirm <= DL_IFI_TIME0); // 组态非法（含 tConfirm 非正与迟滞负值）/ an illegal configuration including a non positive window and a negative hysteresis

// 段 1｜判据预计算与定时器无条件周期刷新（禁入分支，R7）：IN = 三判据合取 AND 使能 AND 无组态故障 / segment 1, the criteria precompute and the unconditional timer refresh
_bFanOk := bFanRun; // 风机运行判据（无迟滞，掉电即失效）/ the fan criterion without hysteresis, it fails as soon as the feedback drops
_bFinSpd := (fAirSpeed = fAirSpeed) AND ((fAirSpeed - fAirSpeed) = (fAirSpeed - fAirSpeed)); // 风速测点有限 / the air speed sample is finite
_bFinBal := (fBalanceV = fBalanceV) AND ((fBalanceV - fBalanceV) = (fBalanceV - fBalanceV)); // 平衡测点有限 / the balance sample is finite
// 迟滞阈值预计算（组态闸在段 2，故此处先按域内假设算，域外值不作为判据依据）/ the hysteresis thresholds are precomputed here, the configuration gate in segment two decides whether they are used
_fPctScale := fHystPct / DL_IFI_HUND; // 迟滞小数化 [−] / the hysteresis as a fraction
_fSpdTrip := fSpeedMin * (1.0 - _fPctScale); // 风速置警阈值 = 下限 × (1 − h) [米每秒] / the trip threshold
_fSpdRele := fSpeedMin * (1.0 + _fPctScale); // 风速复原阈值 = 下限 × (1 + h) [米每秒] / the release threshold
_fBalTrip := fBalanceLimV; // 平衡置警阈值 = 绝对上限 [伏] / the balance trip threshold equals the limit
_fBalRele := fBalanceLimV * (1.0 - _fPctScale); // 平衡复原阈值 = 上限 × (1 − h) [伏] / the balance release threshold
_fBalAbs := ABS(fBalanceV); // 平衡电压绝对值（正负偏等量处理，迟滞对称）[伏] / the absolute balance voltage
// 风速判据：非有限即保守判不满足（边界四）/ the air speed criterion treats a non finite sample as failing
IF _bFinSpd THEN // 测点有限才用迟滞判据 / the hysteresis runs only on a finite sample
    IF NOT _bAlmSpd THEN // 未报警态 / the released state
        IF fAirSpeed < _fSpdTrip THEN // 跌破置警阈值 / below the trip threshold
            _bAlmSpd := TRUE; // 置报警迟滞状态 / set the alarm state
        END_IF
    ELSE // 已报警态 / the tripped state
        IF fAirSpeed > _fSpdRele THEN // 回升超过复原阈值 / above the release threshold
            _bAlmSpd := FALSE; // 复原 / release
        END_IF
    END_IF
    _bSpeedOk := NOT _bAlmSpd; // 判据结果由迟滞状态派生 / the criterion derives from the hysteresis state
ELSE // 测点非有限：保守判不满足并置报警（区分码见段 6）/ a non finite sample conservatively fails and raises the alarm
    _bAlmSpd := TRUE; // 保守落报警态 / conservatively trip
    _bSpeedOk := FALSE; // 判据不满足 / the criterion fails
END_IF
// 平衡判据：非有限即保守判不满足（边界四）/ the balance criterion treats a non finite sample as failing
IF _bFinBal THEN // 测点有限才用迟滞判据 / the hysteresis runs only on a finite sample
    IF NOT _bAlmBal THEN // 未报警态 / the released state
        IF _fBalAbs > _fBalTrip THEN // 超过置警阈值 / above the trip threshold
            _bAlmBal := TRUE; // 置报警迟滞状态 / set the alarm state
        END_IF
    ELSE // 已报警态 / the tripped state
        IF _fBalAbs < _fBalRele THEN // 回落低于复原阈值（限 5 V 时 4.9 V 仍在报警带内）/ below the release threshold, four point nine volts still sits inside the band
            _bAlmBal := FALSE; // 复原 / release
        END_IF
    END_IF
    _bBalOk := NOT _bAlmBal; // 判据结果由迟滞状态派生 / the criterion derives from the hysteresis state
ELSE // 测点非有限：保守判不满足并置报警 / a non finite sample conservatively fails and raises the alarm
    _bAlmBal := TRUE; // 保守落报警态 / conservatively trip
    _bBalOk := FALSE; // 判据不满足 / the criterion fails
END_IF
_bAllOk := _bFanOk AND _bSpeedOk AND _bBalOk; // 三判据合取 / the conjunction
IF _bCfgBad THEN // 组态非法：合取强制失满足（组态阈值不可信，可能是 NaN）/ an illegal configuration forces the conjunction to fail
    _bAllOk := FALSE; // 合取清零（阈值可能是 NaN）/ clear the conjunction, the thresholds may be NaN
END_IF
tonConfirm(IN := _bAllOk AND bEnable AND (NOT _bCfgBad), PT := tConfirm); // 确认窗计时（使能 + 组态闸串入，组态位为本拍值）/ the confirmation window with the enable and the configuration gate in series

// 段 1｜首拍初始化（R310；出厂默认无许可，边界二）/ segment 1, the first scan init with the safe default
IF NOT _bInit THEN // 首拍一拍 / the first scan
    _bInit := TRUE; // 置首拍标志 / raise the first scan flag
    _eState := E_DL_IonFanPhase.eIdle; // 状态显式落空闲 / place the state to idle
    _bAlmSpd := FALSE; // 风速报警迟滞态显式清零 / clear the air speed alarm state explicitly
    _bAlmBal := FALSE; // 平衡报警迟滞态显式清零 / clear the balance alarm state explicitly
    bPermit := FALSE; // 许可显式落假（出厂默认 F）/ force the permit false on the first scan
END_IF

// 段 2｜首拍初始化（R310；出厂默认无许可，边界二）/ segment 2, the first scan init with the safe default
// 段 3｜主状态机（ENUM + CASE，ELSE 兜底并清许可；安全相迁移带全量闸位复检，R274）/ segment 3, the main machine
CASE _eState OF
    E_DL_IonFanPhase.eIdle: // 空闲相（失能时驻留，驻留由分支表达，禁自赋值死语句，R261）/ the idle phase, dwelling is expressed by the branch
        IF bEnable AND _bCfgBad THEN // 使能但组态非法（边界五）/ enabled with an illegal configuration
            _eState := E_DL_IonFanPhase.eAlarm; // 迁入报警相 / enter the alarm phase
        ELSIF bEnable THEN // 使能且组态合法 / enabled with a legal configuration
            _eState := E_DL_IonFanPhase.eWarmup; // 迁入确认相（确认窗自下一拍起计）/ enter the confirmation phase, the window counts from the next scan
        END_IF
    E_DL_IonFanPhase.eWarmup: // 确认相：TON 计时中 / the confirmation phase
        IF (NOT bEnable) OR _bCfgBad THEN // 退出条件一：失能或组态非法（前置条件已消失）/ exit one, the prerequisite disappeared
            _eState := E_DL_IonFanPhase.eAlarm; // 迁入报警相 / enter the alarm phase
        ELSIF tonConfirm.Q AND _bAllOk THEN // 退出条件二：确认窗到且三判据仍满足（安全相迁移全量复检）/ exit two, the window elapsed with the criteria still holding
            _eState := E_DL_IonFanPhase.ePermit; // 迁入已许可相 / enter the permitted phase
        ELSIF NOT _bAllOk THEN // 退出条件三：判据在窗内失效 / exit three, a criterion failed inside the window
            _eState := E_DL_IonFanPhase.eAlarm; // 迁入报警相 / enter the alarm phase
        END_IF
    E_DL_IonFanPhase.ePermit: // 已许可相 / the permitted phase
        IF NOT _bAllOk THEN // 任一判据失效：零延时撤除（边界一）/ any criterion failed, the permit is withdrawn with no delay
            _eState := E_DL_IonFanPhase.eAlarm; // 同拍迁入报警相 / enter the alarm phase on the same scan
        ELSIF (NOT bEnable) OR _bCfgBad THEN // 失能或组态非法 / disabled or an illegal configuration
            _eState := E_DL_IonFanPhase.eAlarm; // 迁入报警相 / enter the alarm phase
        END_IF
    E_DL_IonFanPhase.eAlarm: // 报警相 / the alarm phase
        IF NOT bEnable THEN // 退出条件一：失能 / exit one, disabled
            _eState := E_DL_IonFanPhase.eIdle; // 回空闲 / back to idle
        ELSIF _bAllOk AND (NOT _bCfgBad) THEN // 退出条件二：三判据全恢复且组态合法（须重走确认窗）/ exit two, every criterion recovered, the window restarts
            _eState := E_DL_IonFanPhase.eWarmup; // 回确认相（不直接回许可相，禁跳过确认窗）/ back to confirmation, never jumping straight to permitted
        END_IF
    ELSE // 非法枚举值拦截（边界六：落报警相并清许可，禁静默）/ the illegal enumeration guard
        _eState := E_DL_IonFanPhase.eAlarm; // 落报警相 / force the alarm phase
END_CASE

// 段 4｜统一出口（R191 名实双出口：bPermit 与 eState 同源；安全侧默认 FALSE；三报警位与 bError 全部串 bEnable，v1.0.1 修 R62-D3）/ segment 4, the unified outlet
eState := _eState; // 状态出口 / the state outlet
bPermit := (_eState = E_DL_IonFanPhase.ePermit) AND _bAllOk AND bEnable AND (NOT _bCfgBad); // 许可出口：态 + 合取 + 使能 + 组态四重同源（同拍撤除）/ the permit outlet with four sources, withdrawn on the same scan
bAlarmFan := (NOT bFanRun) AND bEnable; // 风机反馈丧失（Failure 级，无迟滞；串 bEnable，失能不外显假故障，v1.0.1）/ the fan feedback loss without hysteresis, gated by the enable so the disabled phase shows no false failure
bAlarmSpeed := _bAlmSpd AND bEnable; // 风速报警出口（迟滞状态派生；串 bEnable，v1.0.1）/ the air speed alarm outlet gated by the enable
bAlarmBalance := _bAlmBal AND bEnable; // 平衡报警出口（迟滞状态派生；串 bEnable，v1.0.1）/ the balance alarm outlet gated by the enable
bValid := (NOT _bCfgBad) AND _bFinSpd AND _bFinBal; // 测量可用：组态合法且两测点均有限 / usable, a legal configuration and two finite samples
bError := bEnable AND (_bCfgBad OR (NOT _bFinSpd) OR (NOT _bFinBal) OR (NOT bFanRun)); // 故障位串 bEnable（v1.0.1 修 R62-D3：失能相不外显 Failure 级假故障，R45 配对随码回放段同口径）/ the fault bit gated by the enable, aligned with the replay segment

// 段 5｜码位回放（首因保序：组态 → 风机 → 风速测点 → 平衡测点 → 信息级；失能相不发码，v1.0.1）/ segment 5, the code replay with the first cause kept first, silent while disabled
IF NOT bEnable THEN // 失能相：不发任何码（Failure 级假故障不再外显，v1.0.1 修 R62-D3）/ the disabled phase emits no code at all
    eErr := 16#0000_0000; // 归零 / zero
ELSIF _bCfgBad THEN // 组态成因优先 / the configuration cause comes first
    eErr := 16#0003_0717; // 故障级：组态非法 / fault grade, an illegal configuration
ELSIF NOT _bFinSpd THEN // 风速测点坏（与真超标分开，R90）/ the air speed sample is broken, kept apart from a real overshoot
    eErr := 16#0003_0719; // 故障级：风速测点非有限 / fault grade, the air speed sample is not finite
ELSIF NOT _bFinBal THEN // 平衡测点坏 / the balance sample is broken
    eErr := 16#0003_071A; // 故障级：平衡电压测点非有限 / fault grade, the balance sample is not finite
ELSIF NOT bFanRun THEN // 风机反馈丧失（Failure 级）/ the fan feedback loss
    eErr := 16#0003_0718; // 故障级：风机运行反馈丧失 / fault grade, the fan feedback is lost
ELSIF _bAlmSpd THEN // 风速真低于下限（OutOfSpec）/ the air speed really is below the floor
    eErr := 16#0003_071B; // 信息级：风速低于下限 / informational, the air speed is below the floor
ELSIF _bAlmBal THEN // 平衡真超限（OutOfSpec）/ the balance really is over the limit
    eErr := 16#0003_071C; // 信息级：平衡电压超限 / informational, the balance voltage is over the limit
ELSE // 无事件 / no event
    eErr := 16#0000_0000; // 正常 / ok
END_IF
END_FUNCTION_BLOCK

(* ---- FB_DL_LevelSwitchVib.st ---- *)
(*==============================================================================
 * 组件名称 (Component)  : FB_DL_LevelSwitchVib
 * 所属子库 (Sublibrary) : DL_Device
 * 当前版本 (Version)    : 1.0.1
 * 兼容性   (Platform)   : CODESYS 3.5 / TwinCAT 3 / 汇川 InoProShop / Machine Expert
 *                         仅依赖 Standard.library（TON / R_TRIG），零厂商方言
 * 分类     (Category)   : 设备功能块（Function Block，实现 I_DL_LevelSwitch）
 * 功能简述 (Function)   : 振动叉式料位开关信号处理块。原始开关防抖 → 失效安
 *                         全方向归一（fail-safe HIGH/LOW 可选）→ 覆盖/裸露
 *                         双延迟确认 → 有料/无料双联锁输出 + 传感器失效诊
 *                         断镜像（本轮预留）。
 * 接口实现 (Implements) : I_DL_LevelSwitch。接口属性同名成员（eState/bMaterial/
 *                         bHighAlarm/bLowAlarm/bFault/uErrorId）按 R22 以只
 *                         读 PROPERTY GET 承载（内部镜像同源），非接口成员
 *                         bSensorTest 保留 VAR_OUTPUT；方法 CmdReset/CmdTest
 *                         在本文件尾部落地。
 * 公约遵循 (Convention) : 0.1/R23 周期信号处理型（防抖/延迟由 TON 语义承载，
 *                         无初始化/跟踪同步语义），免首扫，无 bInit。
 *                         0.2/R21 bFault 显式排除信息级码；0.5/R7 全部实例
 *                         主体最前部无条件刷新；0.7/R15 故障级锁存仅复位路
 *                         径清码。
 *                         0.8 故障码段位 16#0003_xxxx（经 DL_Device
 *                         VERSION.md 码表核对：规格建议 0003_0290/0003_010a
 *                         中 0290 已由本轮 FB_DL_GuardLockDoor 顺延占用、
 *                         010a 与库内 0110~0116 编号惯例不一致，依公约顺延
 *                         归一）：
 *                         【故障级】0003_02C0 失效安全模式枚举越界；
 *                         【信息级】0003_0116 传感器信号静默提示（预留信息
 *                         级，本轮仅登记码位不触发）。
 * 红线自检 (Redline)    : R1 零全局变量表/外部变量引用 ✓｜R2 零物理 IO 地址 ✓
 *                         R3 纯 IEC 61131-3 ✓｜R4 枚举域防御/参数钳位 ✓
 *                         R5 全变量中英双语同行注释 ✓｜R6 状态映像 IF 派生
 *                         链含 ELSE 兜底（信号处理型派生映像）✓
 *                         R7 四实例（R_TRIG×1/TON×4）主体最前部无条件刷新 ✓
 *                         R8 全常量化 ✓
 * 设计要点 (Key notes)  : ① 失效安全归一核心：bMaterial 归一式 bRawSwitch
 *                           XOR (eFailSafeMode = eLow) 的语义等价式（用 IF
 *                           显式写，禁 XOR 技巧裸用）——eHigh 组态下原始信
 *                           号直接作为有料判定；eLow 组态约定传感器原始信号
 *                           极性为 TRUE=无料/裸露（出厂反相接线，接线层保
 *                           证），取反后统一为 TRUE=有料，防现场接反；
 *                         ② bEnable=FALSE 或传感器失效时输出强制归一到安全
 *                           侧：eHigh → 强制有料（bHighAlarm 报警，防溢流）；
 *                           eLow → 强制无料（bLowAlarm 报警，防干转）；
 *                         ③ 高/低联锁方向语义写死：bHighAlarm = 归一后有料
 *                           （eHigh 失效即报警）；bLowAlarm = 归一后无料
 *                           （eLow 失效即报警），两输出方向由本归一约定承
 *                           载，现场不得反接；
 *                         ④ 覆盖/裸露双延迟：防抖 TON×2 + 确认 TON×2 全部
 *                           在主体前部无条件刷新（R7）；
 *                         ⑤ 传感器失效检测（信号静默）本轮预留：码位
 *                           0003_0116 与 eSensorLoss 态已登记，检测算法后续
 *                           轮次落地（R11 留档）。
 * 偏离留档 (Deviation)  : 依 R11 头注释留档，共 1 条：
 *                         ① 码位顺延归一：规格建议 0003_0290 与本轮
 *                           FB_DL_GuardLockDoor 顺延占用冲突，取 0003_02C0；
 *                           规格建议 0003_010a 改为 0003_0116 与库内信息级
 *                           编号惯例一致（核对结果优先于建议值）。
 * 开源溯源 (Origin)     : 来源标签 tcopen-component / level-switch-failsafe
 *                         （RAW_NOTES_R7 S-7：TcOpen 料位开关组件失效安全
 *                         语义域与振动叉开关防抖/双延迟公开惯例，公开资料，
 *                         仅借鉴语义域；归一实现、码位与引脚契约 100% 本库
 *                         独立设计，clean-room 未复制源码）。
 * 验收向量 (Acceptance) :
 *   V1 有料/无料双延迟切换逐拍：raw 稳定翻转 → tDebounce 过 → tCoverDelay/
 *      tBareDelay 过 → bMaterial 翻转；
 *   V2 fail-safe HIGH 断线注入（使能切断模拟失效）：bEnable=FALSE + eHigh →
 *      bMaterial 强制 TRUE、bHighAlarm=TRUE（防溢流方向）；
 *   V3 fail-safe LOW 断线注入：bEnable=FALSE + eLow → bMaterial 强制 FALSE、
 *      bLowAlarm=TRUE（防干转方向）；
 *   V4 模式枚举越界：eFailSafeMode 写入域外值 → 故障锁存 0003_02C0；
 *   V5 复位：bReset 沿 → 故障清零回 eIdle 镜像态。
 * 修订历史 (Revision)   :
 *   2026-11-15  v1.0.0  首版入库（Round 07 · DL_Device 料位开关族实现件）
 *   2026-11-15  v1.0.1  终审修复 1 处：_fbTrigTest 误接 bEnable——每次使能
 *                       上升沿（含正常开机）误置 bSensorTest 测试镜像一拍，
 *                       删除误接实例，bSensorTest 仅由 CmdTest 单拍承载
 *============================================================================*)
FUNCTION_BLOCK FB_DL_LevelSwitchVib IMPLEMENTS I_DL_LevelSwitch
VAR_INPUT
    bRawSwitch    : BOOL;               // 传感器原始开关信号（Raw switch signal），TRUE=触点动作（介质覆盖叉体，按传感器极性定义）/ Raw switch, TRUE = contact acted per sensor polarity
    eFailSafeMode : E_DL_FailSafeMode := E_DL_FailSafeMode.eHigh; // 失效安全模式（Fail-safe mode），eHigh=失效报有料（防溢流）/ eLow=失效报无料（防干转）/ Fail-safe direction
    tDebounce     : TIME := T#200MS;    // 防抖窗口（Debounce），默认 T#200MS / Debounce window
    tCoverDelay   : TIME := T#1S;       // 覆盖确认延迟（Cover delay），默认 T#1S，防液面波动误翻转 / Cover confirm delay
    tBareDelay    : TIME := T#1S;       // 裸露确认延迟（Bare delay），默认 T#1S / Bare confirm delay
    bEnable       : BOOL;               // 处理使能（Processing enable），FALSE=输出按失效安全方向强制镜像 / FALSE forces fail-safe mirrored outputs
    bReset        : BOOL;               // 上升沿复位故障（Reset edge）/ Rising edge resets fault
END_VAR
VAR_OUTPUT
    bSensorTest : BOOL;                 // 传感器测试态镜像（Sensor test mirror），CmdTest 期间一拍 / Test mirror, one scan during CmdTest
END_VAR
VAR
    _eState        : E_DL_LevelState;   // 派生诊断状态（Derived diagnostic state），属性只读 / Derived state, read-only via property
    _bFaultLatch   : BOOL;              // 故障锁存标志（Fault latch flag），仅复位路径清除 / Fault latch, cleared only via reset path
    _uErrorIdInt   : UDINT;             // 内部故障级码寄存（Internal fault-level register）/ Internal fault-level register
    _uInfoCode     : UDINT;             // 本拍信息级码（Info code this cycle），瞬时型每拍重算 / Transient info code, recomputed each scan
    _bModeValid    : BOOL;              // 失效安全模式枚举合法（Fail-safe mode in domain）/ Mode in-domain flag
    _bRawDebounced : BOOL;              // 防抖后原始信号（Debounced raw signal）/ Debounced raw signal
    _bMatNorm      : BOOL;              // 极性归一后有料判定（Polarity-normalized material）/ Polarity-normalized material
    _bMatSafe      : BOOL;              // 失效安全归一输出（Fail-safe normalized material output）/ Fail-safe normalized output
    _bMatConfirmed : BOOL;              // 双延迟确认后有料判定（Delay-confirmed material）/ Delay-confirmed material
    _bTestPulse    : BOOL;              // 测试态单拍请求（Test one-shot request）/ Test one-shot request
    _bPendReset    : BOOL;              // 方法复位请求（Method reset request）/ Method reset request
    _bPendTest     : BOOL;              // 方法测试请求（Method test request）/ Method test request
    _fbTrigReset   : R_TRIG;            // 引脚复位沿（Pin reset edge）/ Pin reset edge detector
    _fbTonDbCover  : TON;               // 原始信号覆盖侧防抖（Raw cover-side debounce）/ Cover-side debounce timer
    _fbTonDbBare   : TON;               // 原始信号裸露侧防抖（Raw bare-side debounce）/ Bare-side debounce timer
    _fbTonCover    : TON;               // 覆盖确认延迟（Cover confirm delay）/ Cover confirm delay
    _fbTonBare     : TON;               // 裸露确认延迟（Bare confirm delay）/ Bare confirm delay
END_VAR

METHOD CmdReset : BOOL
VAR_INPUT
END_VAR
IF _bFaultLatch OR (_eState = E_DL_LevelState.eFault) THEN
    _bPendReset := TRUE;          // 登记复位请求（Register reset request）
    CmdReset := TRUE;             // 可复位（Resettable）
ELSE
    CmdReset := FALSE;            // 无故障可复位（Nothing to reset）
END_IF

(*------------------------------------------------------------------------------
 * 方法: CmdTest —— 传感器功能测试请求：输出镜像进入测试态一拍。故障态拒绝。
 *      Method CmdTest - sensor test request, test mirror one scan, rejected in fault.
 *------------------------------------------------------------------------------*)
    END_METHOD

METHOD CmdTest : BOOL
VAR_INPUT
END_VAR
IF _bFaultLatch OR (_eState = E_DL_LevelState.eFault) THEN
    CmdTest := FALSE;             // 故障态拒绝（Rejected in fault）
ELSE
    _bPendTest := TRUE;           // 登记测试请求（Register test request）
    CmdTest := TRUE;              // 受理成功（Accepted）
END_IF

(*------------------------------------------------------------------------------
 * 属性: eState（GET）—— 当前诊断状态只读视图。
 *      Property eState (GET) - read-only diagnostic state view.
 *------------------------------------------------------------------------------*)
    END_METHOD

// ============================================================================
// 段 1｜实例无条件周期刷新（R7/0.5：严禁置于 IF/CASE 分支内）
//      Unconditional per-cycle refresh of all instances (R7/0.5)
// ============================================================================
_fbTrigReset(CLK := bReset);
_fbTonDbCover(IN := bRawSwitch, PT := tDebounce);           // 覆盖侧防抖（Cover debounce）
_fbTonDbBare(IN := (NOT bRawSwitch), PT := tDebounce);      // 裸露侧防抖（Bare debounce）
_fbTonCover(IN := _bRawDebounced AND (NOT _bMatConfirmed) AND (NOT _bFaultLatch), PT := tCoverDelay); // 覆盖确认（Cover confirm）
_fbTonBare(IN := (NOT _bRawDebounced) AND _bMatConfirmed AND (NOT _bFaultLatch), PT := tBareDelay);   // 裸露确认（Bare confirm）

// ============================================================================
// 段 2｜模式域防御 + 信息级预清零 + 复位路径（R15）
//      Mode domain guard + info preset + reset path (R15)
// ============================================================================
_uInfoCode := 0;                  // 信息级瞬时型每拍重算（Transient info recomputed each scan）
_bModeValid := (eFailSafeMode = E_DL_FailSafeMode.eHigh) OR (eFailSafeMode = E_DL_FailSafeMode.eLow); // 模式域校验（Mode domain check）
IF NOT _bModeValid THEN
    _bFaultLatch := TRUE;         // 模式枚举越界锁存（Mode out-of-domain latch）
    _uErrorIdInt := 16#0003_02C0; // 0003_02C0 失效安全模式枚举越界【故障级】/ Fail-safe mode out of domain, fault level
END_IF

IF _fbTrigReset.Q OR _bPendReset THEN
    _bPendReset := FALSE;         // 消费方法复位请求（Consume method reset）
    IF _bModeValid THEN           // 故障源已消失才解除（Release only when source gone）
        _bFaultLatch := FALSE;    // 故障锁存解除（Fault latch released）
        _uErrorIdInt := 16#0000_0000; // 故障码清零（Fault code cleared）
    END_IF
END_IF

// ============================================================================
// 段 3｜防抖合成 + 失效安全归一（核心语义，IF 显式写，禁 XOR 裸用）
//      Debounce merge + fail-safe normalization (explicit IF, no raw XOR)
// ============================================================================
IF _fbTonDbCover.Q THEN
    _bRawDebounced := TRUE;       // 覆盖侧防抖达成（Cover debounce reached）
ELSIF _fbTonDbBare.Q THEN
    _bRawDebounced := FALSE;      // 裸露侧防抖达成（Bare debounce reached）
END_IF                            // 窗内保持上次判定（Hold previous verdict inside window）

IF NOT _bModeValid THEN
    _bMatNorm := FALSE;           // 模式非法归一安全侧（Invalid mode normalized to safe side）
ELSIF eFailSafeMode = E_DL_FailSafeMode.eLow THEN
    _bMatNorm := NOT _bRawDebounced; // eLow 极性取反归一（约定 raw TRUE=无料/裸露，反相接线层保证）/ eLow polarity inversion (raw TRUE = bare by wiring convention)
ELSE
    _bMatNorm := _bRawDebounced;  // eHigh 极性直通归一（raw TRUE=覆盖有料）/ eHigh polarity pass-through
END_IF

// 使能切断/故障期强制镜像到失效安全侧（eHigh→有料防溢流；eLow→无料防干转）
// Enable-off or fault forces the fail-safe side (eHigh → covered, eLow → bare)
IF (NOT bEnable) OR _bFaultLatch THEN
    IF eFailSafeMode = E_DL_FailSafeMode.eHigh THEN
        _bMatSafe := TRUE;        // eHigh 强制有料（Force covered, overflow-safe）
    ELSE
        _bMatSafe := FALSE;       // eLow 强制无料（Force bare, dry-run-safe）
    END_IF
ELSE
    _bMatSafe := _bMatNorm;       // 正常处理直通（Normal processing pass-through）
END_IF

// ============================================================================
// 段 4｜覆盖/裸露双延迟确认 + 测试单拍 + 状态映像（IF 派生链含 ELSE 兜底）
//      Cover/bare dual-delay confirm + test one-shot + state image with ELSE
// ============================================================================
IF _fbTonCover.Q THEN
    _bMatConfirmed := TRUE;       // 覆盖确认达成（Cover confirmed）
ELSIF _fbTonBare.Q THEN
    _bMatConfirmed := FALSE;      // 裸露确认达成（Bare confirmed）
END_IF                            // 确认窗内保持（Hold inside confirm window）

IF _bFaultLatch THEN
    _eState := E_DL_LevelState.eFault;      // 故障映像（Fault image）
ELSIF (NOT bEnable) THEN
    _eState := E_DL_LevelState.eSensorLoss; // 使能切断：失效安全强制镜像的诊断映像（强制镜像诊断位）/ Enable-off: forced-mirror diagnostic image
ELSIF _bMatConfirmed THEN
    _eState := E_DL_LevelState.eMaterial;   // 有料确认映像（Material image）
ELSE
    _eState := E_DL_LevelState.eNoMaterial; // 无料兜底映像（No-material fallback image）
END_IF

bSensorTest := _bPendTest;        // 测试态镜像一拍，仅由 CmdTest 承载（v1.0.1 修复：原
                                  // _fbTrigTest 误接 bEnable，使能沿误置测试镜像）
                                  // Test mirror one scan, CmdTest only (v1.0.1 fix)
_bPendTest := FALSE;              // 方法测试请求消费（Method test request consumed）

(*------------------------------------------------------------------------------
 * 方法: CmdReset —— 复位故障。仅故障态受理（接口方法拒绝语义红线）。
 *      Method CmdReset - reset, accepted only in fault state.
 *------------------------------------------------------------------------------*)

PROPERTY eState : E_DL_LevelState
eState := _eState;                // 返回派生状态（Return derived state）

(*------------------------------------------------------------------------------
 * 属性: bMaterial（GET）—— 有料判定输出（失效安全归一后，TRUE=有料）。
 *      Property bMaterial (GET) - fail-safe normalized material output.
 *------------------------------------------------------------------------------*)
PROPERTY bMaterial : BOOL
bMaterial := _bMatSafe;           // 返回失效安全归一输出（Return fail-safe normalized output）

(*------------------------------------------------------------------------------
 * 属性: bHighAlarm（GET）—— 高点溢流联锁输出（fail-safe HIGH 语义：归一有
 *         料即报警；eHigh 组态下失效即报警，防溢流方向，现场不得反接）。
 *      Property bHighAlarm (GET) - high-level interlock, fail-safe HIGH semantics.
 *------------------------------------------------------------------------------*)
PROPERTY bHighAlarm : BOOL
bHighAlarm := _bMatSafe;          // 有料即高点报警（Covered = high alarm）

(*------------------------------------------------------------------------------
 * 属性: bLowAlarm（GET）—— 低点干转联锁输出（fail-safe LOW 语义：归一无料
 *         即报警；eLow 组态下失效即报警，防干转方向，现场不得反接）。
 *      Property bLowAlarm (GET) - low-level interlock, fail-safe LOW semantics.
 *------------------------------------------------------------------------------*)
PROPERTY bLowAlarm : BOOL
bLowAlarm := NOT _bMatSafe;       // 无料即低点报警（Bare = low alarm）

(*------------------------------------------------------------------------------
 * 属性: bFault（GET）—— 故障锁存指示（信息级码不置本位，0.2 公约）。
 *      Property bFault (GET) - fault latch indicator, info codes excluded.
 *------------------------------------------------------------------------------*)
PROPERTY bFault : BOOL
bFault := _bFaultLatch OR (_eState = E_DL_LevelState.eFault); // 显式排除信息级派生式（Derived form excluding info codes）

(*------------------------------------------------------------------------------
 * 属性: uErrorId（GET）—— 末次故障码（故障级优先，无故障时透出本拍信息级
 *         码，0.2/0.15 公约；0003_0116 为预留信息级，本轮不触发）。
 *      Property uErrorId (GET) - last error code (fault priority, info shown otherwise).
 *------------------------------------------------------------------------------*)
PROPERTY uErrorId : UDINT
IF (_uErrorIdInt <> 0) OR (_eState = E_DL_LevelState.eFault) THEN
    uErrorId := _uErrorIdInt;     // 故障级码优先透出（Fault-level priority）
ELSE
    uErrorId := _uInfoCode;       // 无故障时透出本拍信息级码（Transient info code）
END_IF
END_FUNCTION_BLOCK
